(* IEC 61131-3 sources: llm-plc-st-eval/data/processed_definitivo/qwen2.5-coder_14b/B8/few_shot, 3 files *)

(* ---- ejec_1.st ---- *)
FUNCTION_BLOCK FB_Puerta
VAR_INPUT
    puertaAbierta : BOOL; (* Señal de puerta abierta *)
    reset : BOOL; (* Botón de reset *)
END_VAR
VAR_OUTPUT
    aviso : BOOL; (* Salida de aviso *)
    nAperturas : INT; (* Número de aperturas *)
END_VAR
VAR
    puertaAbiertaAnterior : BOOL; (* Estado anterior de la puerta *)
END_VAR

(* Reinicio del registro *)
IF reset THEN
    nAperturas := 0;
    aviso := FALSE;
END_IF

(* Detección de transición de FALSE a TRUE *)
IF puertaAbierta AND NOT puertaAbiertaAnterior THEN
    nAperturas := nAperturas + 1;
END_IF

(* Actualización del estado anterior *)
puertaAbiertaAnterior := puertaAbierta;

(* Activación del aviso si se alcanzan 5 aperturas *)
IF nAperturas >= 5 THEN
    aviso := TRUE;
END_IF
END_FUNCTION_BLOCK

(* ---- ejec_2.st ---- *)
FUNCTION_BLOCK FB_Puerta
VAR_INPUT
    puertaAbierta : BOOL; (* Señal de puerta abierta *)
    reset : BOOL; (* Botón de reinicio *)
END_VAR
VAR_OUTPUT
    aviso : BOOL; (* Salida de aviso *)
    nAperturas : INT; (* Contador de aperturas *)
END_VAR
VAR
    puertaAbiertaAnterior : BOOL; (* Estado anterior de la puerta *)
END_VAR

(* Reinicio del contador y aviso *)
IF reset THEN
    nAperturas := 0;
    aviso := FALSE;
ELSE
    (* Detección de transición de FALSE a TRUE *)
    IF NOT puertaAbiertaAnterior AND puertaAbierta THEN
        nAperturas := nAperturas + 1;
    END_IF

    (* Activación del aviso si se alcanzan 5 aperturas *)
    aviso := nAperturas >= 5;
END_IF

(* Actualización del estado anterior de la puerta *)
puertaAbiertaAnterior := puertaAbierta;
END_FUNCTION_BLOCK

(* ---- ejec_3.st ---- *)
FUNCTION_BLOCK FB_Puerta
VAR_INPUT
    puertaAbierta : BOOL; (* Señal de puerta abierta *)
    reset : BOOL; (* Botón de reset *)
END_VAR
VAR_OUTPUT
    aviso : BOOL; (* Salida de aviso *)
    nAperturas : INT; (* Número de aperturas *)
END_VAR
VAR
    puertaAbiertaAnterior : BOOL; (* Estado anterior de la puerta abierta *)
END_VAR

(* Reinicio del registro *)
IF reset THEN
    nAperturas := 0;
    aviso := FALSE;
ELSE
    (* Detección de transición de FALSE a TRUE *)
    IF NOT puertaAbiertaAnterior AND puertaAbierta THEN
        nAperturas := nAperturas + 1;
    END_IF

    (* Activación del aviso si se alcanzan 5 aperturas *)
    aviso := nAperturas >= 5;
END_IF

(* Actualización del estado anterior de la puerta *)
puertaAbiertaAnterior := puertaAbierta;
END_FUNCTION_BLOCK
